// TIA Portal V15.1 export
// export: Created 2026-11-02T18:55:10.9093708Z, ExportSetting WithDefaults, DisplayName Totally Integrated Automation Portal, DisplayVersion V15.1, DisplayName TIA Portal Openness, DisplayVersion V15.1, DisplayName STEP 7 Professional, DisplayVersion V15.1, DisplayName WinCC Professional, DisplayVersion V15.1
FUNCTION_BLOCK "Scrubber"   // FB2, LAD
TITLE = Scrubber
{ S7_Optimized_Access := 'TRUE' }
VERSION : 0.1
// Gas scrubber, docs/التشغيل.md §1
// stored: AutoNumber false, IsIECCheckEnabled false, IsRetainMemResEnabled false, MemoryReserve 100, SetENOAutomatically False, UDAEnableTagReadback false
   VAR_INPUT
      PSH : Bool;   // PSH-101 healthy (contact closed)
      LSH : Bool;   // LSH-102 healthy
      LSHH : Bool;   // LSHH-103 healthy
      EStopOK : Bool;   // Sys.EStopOK
      ResetPulse : Bool;   // Sys.ResetPulse
      FirstScan : Bool;   // Sys.FirstScan
      TDrnOn : Time;   // Par.TDrnOn_V (C04)
      TDrnOff : Time;   // Par.TDrnOff_V (C04)
      TDrnMax : Time;   // Par.TDrnMax_V (C04a)
   END_VAR
   VAR_OUTPUT
      Tripped : Bool;   // Suction trip latch C01/C02/C03/C05: XV-403 closed until RESET
      FlareTrip : Bool;   // Flare trip latch C01/C02/C03: XV-401 open until RESET
      ValvesNormal : Bool;   // No trip latched: flare closed and suction open (HMI)
      FlareCmd : Bool;   // Q0.2 XV-401 (NO): 1 = energised = closed
      DrainCmd : Bool;   // Q0.3 XV-402 (NC): 1 = energised = open (C04 / C05)
      SuctionCmd : Bool;   // Q0.4 XV-403 (NC): 1 = energised = open
      F_DrainTO : Bool;   // C04a: drain open too long, latched until RESET
      F_LshFault : Bool;   // C04b: LSHH-103 without LSH-102, latched until RESET
      Alm_PSH : Bool;   // HMI alarm C03
      Alm_LSH : Bool;   // HMI alarm C04
      Alm_LSHH : Bool;   // HMI alarm C05
      Cause_EStop : Bool;   // C06a / F44: E-STOP cause, latched until healthy RESET
      Cause_PSH : Bool;   // C06a / F44: PSH-101 cause, latched until healthy RESET
      Cause_LSHH : Bool;   // C06a / F44: LSHH-103 cause, latched until healthy RESET
      Cause_PwrUp : Bool;   // C06a / F44: power-up cause, latched until healthy RESET
      FirstOut : Int;   // C06a / 0007 D5: 0 none, 1 E-STOP, 2 PSH, 3 LSHH, 4 power-up
   END_VAR
   VAR
      LevelHigh : Bool;
      DrnDemand : Bool;
      T_DrnOn : TON_TIME;
      T_DrnOff : TON_TIME;
      T_DrnMax : TON_TIME;
      T_LshFlt : TON_TIME;
   END_VAR
BEGIN

REGION Network 1: C04 — LSH-102 high level alarm
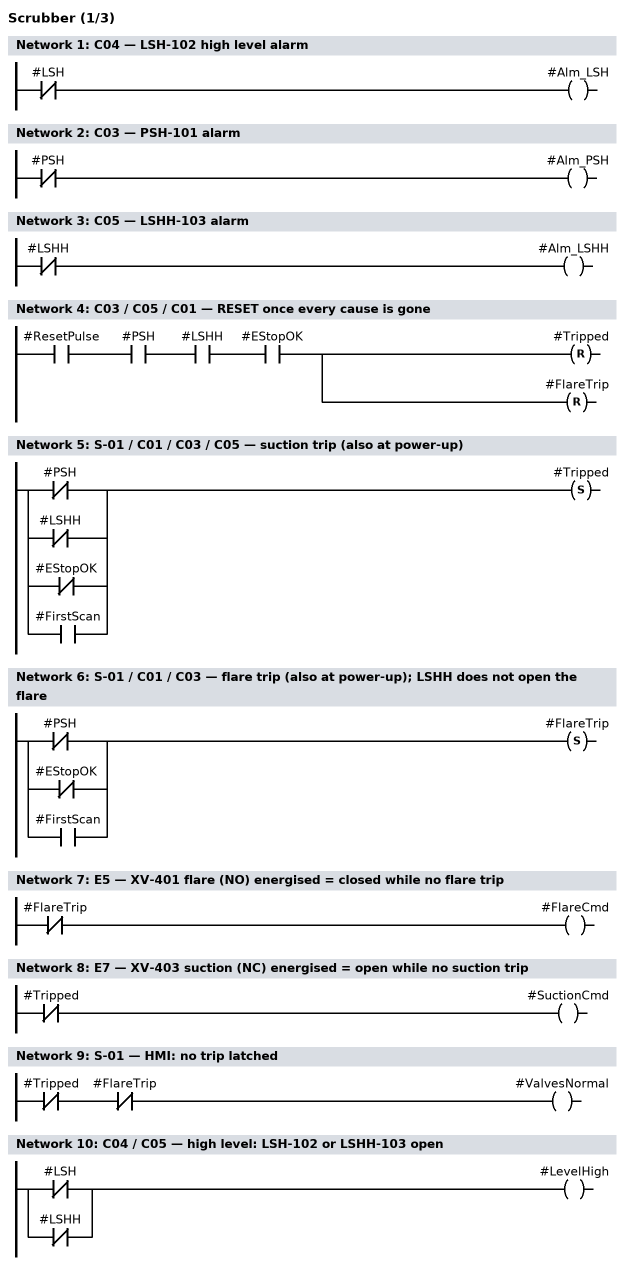
   RUNG wire#powerrail
      I_Contact( #LSH )
      Coil( #Alm_LSH )
   END_RUNG
   // the same network as SCL:
   #Alm_LSH := NOT #LSH;
END_REGION

REGION Network 2: C03 — PSH-101 alarm
   RUNG wire#powerrail
      I_Contact( #PSH )
      Coil( #Alm_PSH )
   END_RUNG
   // the same network as SCL:
   #Alm_PSH := NOT #PSH;
END_REGION

REGION Network 3: C05 — LSHH-103 alarm
   RUNG wire#powerrail
      I_Contact( #LSHH )
      Coil( #Alm_LSHH )
   END_RUNG
   // the same network as SCL:
   #Alm_LSHH := NOT #LSHH;
END_REGION

REGION Network 4: C03 / C05 / C01 — RESET once every cause is gone
   RUNG wire#powerrail
      Contact( #ResetPulse )
      Contact( #PSH )
      Contact( #LSHH )
      Contact( #EStopOK )
      wire#w1
      R_Coil( #Tripped )
   END_RUNG
   RUNG wire#w1
      R_Coil( #FlareTrip )
   END_RUNG
   // the same network as SCL:
   IF #ResetPulse AND #PSH AND #LSHH AND #EStopOK THEN
       #Tripped := FALSE;
       #FlareTrip := FALSE;
   END_IF;
END_REGION

REGION Network 5: S-01 / C01 / C03 / C05 — suction trip (also at power-up)
   RUNG wire#powerrail
      I_Contact( #PSH )
      wire#w1
      S_Coil( #Tripped )
   END_RUNG
   RUNG wire#powerrail
      I_Contact( #LSHH )
   END_RUNG wire#w1
   RUNG wire#powerrail
      I_Contact( #EStopOK )
   END_RUNG wire#w1
   RUNG wire#powerrail
      Contact( #FirstScan )
   END_RUNG wire#w1
   // the same network as SCL:
   IF NOT #PSH OR NOT #LSHH OR NOT #EStopOK OR #FirstScan THEN #Tripped := TRUE; END_IF;
END_REGION

REGION Network 6: S-01 / C01 / C03 — flare trip (also at power-up); LSHH does not open the flare
   RUNG wire#powerrail
      I_Contact( #PSH )
      wire#w1
      S_Coil( #FlareTrip )
   END_RUNG
   RUNG wire#powerrail
      I_Contact( #EStopOK )
   END_RUNG wire#w1
   RUNG wire#powerrail
      Contact( #FirstScan )
   END_RUNG wire#w1
   // the same network as SCL:
   IF NOT #PSH OR NOT #EStopOK OR #FirstScan THEN #FlareTrip := TRUE; END_IF;
END_REGION

REGION Network 7: E5 — XV-401 flare (NO) energised = closed while no flare trip
   RUNG wire#powerrail
      I_Contact( #FlareTrip )
      Coil( #FlareCmd )
   END_RUNG
   // the same network as SCL:
   #FlareCmd := NOT #FlareTrip;
END_REGION

REGION Network 8: E7 — XV-403 suction (NC) energised = open while no suction trip
   RUNG wire#powerrail
      I_Contact( #Tripped )
      Coil( #SuctionCmd )
   END_RUNG
   // the same network as SCL:
   #SuctionCmd := NOT #Tripped;
END_REGION

REGION Network 9: S-01 — HMI: no trip latched
   RUNG wire#powerrail
      I_Contact( #Tripped )
      I_Contact( #FlareTrip )
      Coil( #ValvesNormal )
   END_RUNG
   // the same network as SCL:
   #ValvesNormal := NOT #Tripped AND NOT #FlareTrip;
END_REGION

REGION Network 10: C04 / C05 — high level: LSH-102 or LSHH-103 open
   RUNG wire#powerrail
      I_Contact( #LSH )
      wire#w1
      Coil( #LevelHigh )
   END_RUNG
   RUNG wire#powerrail
      I_Contact( #LSHH )
   END_RUNG wire#w1
   // the same network as SCL:
   #LevelHigh := NOT #LSH OR NOT #LSHH;
END_REGION

REGION Network 11: C04 — drain demand after TDRN_ON of high level
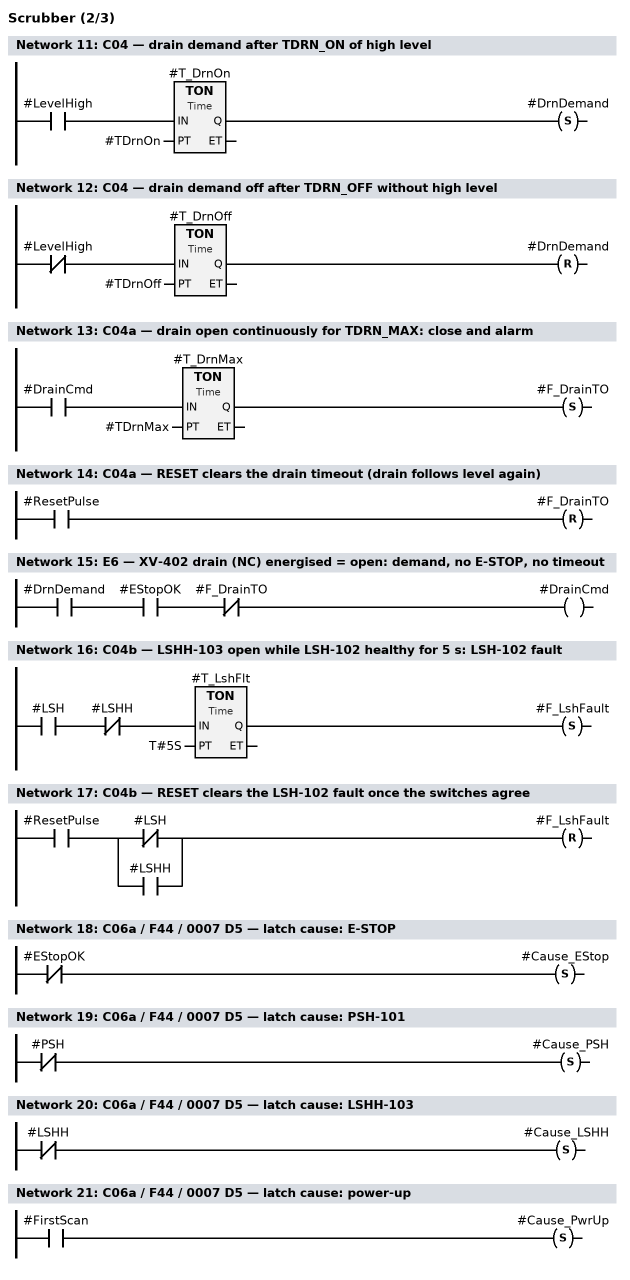
   RUNG wire#powerrail
      Contact( #LevelHigh )
      { S7_Templates := "time_type := Time" } #T_DrnOn.TON(pt := #TDrnOn, et =>)
      S_Coil( #DrnDemand )
   END_RUNG
   // the same network as SCL:
   #T_DrnOn(IN := #LevelHigh, PT := #TDrnOn);   // TON
   IF #T_DrnOn.Q THEN #DrnDemand := TRUE; END_IF;
END_REGION

REGION Network 12: C04 — drain demand off after TDRN_OFF without high level
   RUNG wire#powerrail
      I_Contact( #LevelHigh )
      { S7_Templates := "time_type := Time" } #T_DrnOff.TON(pt := #TDrnOff, et =>)
      R_Coil( #DrnDemand )
   END_RUNG
   // the same network as SCL:
   #T_DrnOff(IN := NOT #LevelHigh, PT := #TDrnOff);   // TON
   IF #T_DrnOff.Q THEN #DrnDemand := FALSE; END_IF;
END_REGION

REGION Network 13: C04a — drain open continuously for TDRN_MAX: close and alarm
   RUNG wire#powerrail
      Contact( #DrainCmd )
      { S7_Templates := "time_type := Time" } #T_DrnMax.TON(pt := #TDrnMax, et =>)
      S_Coil( #F_DrainTO )
   END_RUNG
   // the same network as SCL:
   #T_DrnMax(IN := #DrainCmd, PT := #TDrnMax);   // TON
   IF #T_DrnMax.Q THEN #F_DrainTO := TRUE; END_IF;
END_REGION

REGION Network 14: C04a — RESET clears the drain timeout (drain follows level again)
   RUNG wire#powerrail
      Contact( #ResetPulse )
      R_Coil( #F_DrainTO )
   END_RUNG
   // the same network as SCL:
   IF #ResetPulse THEN #F_DrainTO := FALSE; END_IF;
END_REGION

REGION Network 15: E6 — XV-402 drain (NC) energised = open: demand, no E-STOP, no timeout
   RUNG wire#powerrail
      Contact( #DrnDemand )
      Contact( #EStopOK )
      I_Contact( #F_DrainTO )
      Coil( #DrainCmd )
   END_RUNG
   // the same network as SCL:
   #DrainCmd := #DrnDemand AND #EStopOK AND NOT #F_DrainTO;
END_REGION

REGION Network 16: C04b — LSHH-103 open while LSH-102 healthy for 5 s: LSH-102 fault
   RUNG wire#powerrail
      Contact( #LSH )
      I_Contact( #LSHH )
      { S7_Templates := "time_type := Time" } #T_LshFlt.TON(pt := T#5S, et =>)
      S_Coil( #F_LshFault )
   END_RUNG
   // the same network as SCL:
   #T_LshFlt(IN := #LSH AND NOT #LSHH, PT := T#5S);   // TON
   IF #T_LshFlt.Q THEN #F_LshFault := TRUE; END_IF;
END_REGION

REGION Network 17: C04b — RESET clears the LSH-102 fault once the switches agree
   RUNG wire#powerrail
      Contact( #ResetPulse )
      wire#w1
      I_Contact( #LSH )
      wire#w2
      R_Coil( #F_LshFault )
   END_RUNG
   RUNG wire#w1
      Contact( #LSHH )
   END_RUNG wire#w2
   // the same network as SCL:
   IF #ResetPulse AND (NOT #LSH OR #LSHH) THEN #F_LshFault := FALSE; END_IF;
END_REGION

REGION Network 18: C06a / F44 / 0007 D5 — latch cause: E-STOP
   RUNG wire#powerrail
      I_Contact( #EStopOK )
      S_Coil( #Cause_EStop )
   END_RUNG
   // the same network as SCL:
   IF NOT #EStopOK THEN #Cause_EStop := TRUE; END_IF;
END_REGION

REGION Network 19: C06a / F44 / 0007 D5 — latch cause: PSH-101
   RUNG wire#powerrail
      I_Contact( #PSH )
      S_Coil( #Cause_PSH )
   END_RUNG
   // the same network as SCL:
   IF NOT #PSH THEN #Cause_PSH := TRUE; END_IF;
END_REGION

REGION Network 20: C06a / F44 / 0007 D5 — latch cause: LSHH-103
   RUNG wire#powerrail
      I_Contact( #LSHH )
      S_Coil( #Cause_LSHH )
   END_RUNG
   // the same network as SCL:
   IF NOT #LSHH THEN #Cause_LSHH := TRUE; END_IF;
END_REGION

REGION Network 21: C06a / F44 / 0007 D5 — latch cause: power-up
   RUNG wire#powerrail
      Contact( #FirstScan )
      S_Coil( #Cause_PwrUp )
   END_RUNG
   // the same network as SCL:
   IF #FirstScan THEN #Cause_PwrUp := TRUE; END_IF;
END_REGION

REGION Network 22: C06a / F44 / 0007 D5 — first-out 1: E-STOP (only if none)
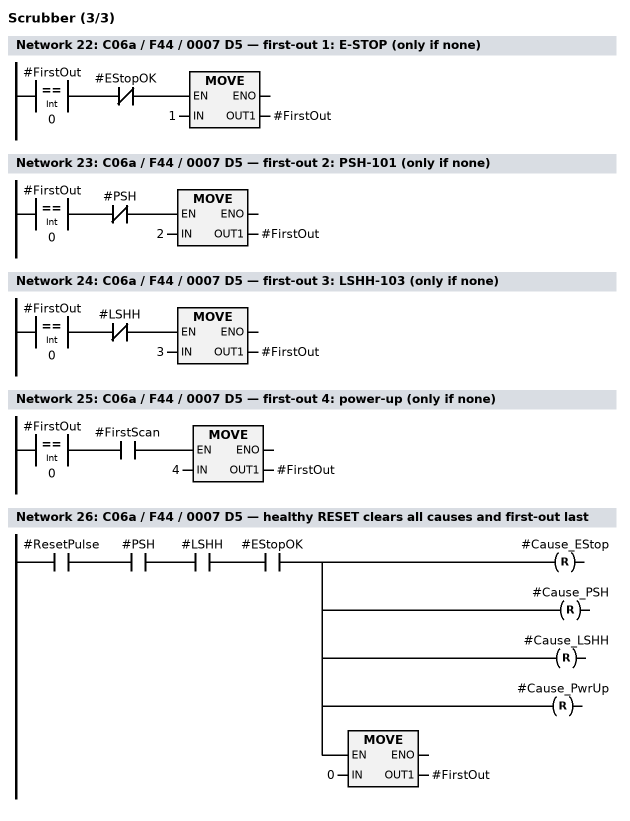
   RUNG wire#powerrail
      { S7_Templates := "SrcType := Int" } EQ_Contact(in1 := #FirstOut, in2 := 0)
      I_Contact( #EStopOK )
      { S7_GenerateENO := "TRUE" } Move(in := 1, out1 => #FirstOut)
   END_RUNG
   // the same network as SCL:
   IF (#FirstOut = 0) AND NOT #EStopOK THEN #FirstOut := 1; END_IF;
END_REGION

REGION Network 23: C06a / F44 / 0007 D5 — first-out 2: PSH-101 (only if none)
   RUNG wire#powerrail
      { S7_Templates := "SrcType := Int" } EQ_Contact(in1 := #FirstOut, in2 := 0)
      I_Contact( #PSH )
      { S7_GenerateENO := "TRUE" } Move(in := 2, out1 => #FirstOut)
   END_RUNG
   // the same network as SCL:
   IF (#FirstOut = 0) AND NOT #PSH THEN #FirstOut := 2; END_IF;
END_REGION

REGION Network 24: C06a / F44 / 0007 D5 — first-out 3: LSHH-103 (only if none)
   RUNG wire#powerrail
      { S7_Templates := "SrcType := Int" } EQ_Contact(in1 := #FirstOut, in2 := 0)
      I_Contact( #LSHH )
      { S7_GenerateENO := "TRUE" } Move(in := 3, out1 => #FirstOut)
   END_RUNG
   // the same network as SCL:
   IF (#FirstOut = 0) AND NOT #LSHH THEN #FirstOut := 3; END_IF;
END_REGION

REGION Network 25: C06a / F44 / 0007 D5 — first-out 4: power-up (only if none)
   RUNG wire#powerrail
      { S7_Templates := "SrcType := Int" } EQ_Contact(in1 := #FirstOut, in2 := 0)
      Contact( #FirstScan )
      { S7_GenerateENO := "TRUE" } Move(in := 4, out1 => #FirstOut)
   END_RUNG
   // the same network as SCL:
   IF (#FirstOut = 0) AND #FirstScan THEN #FirstOut := 4; END_IF;
END_REGION

REGION Network 26: C06a / F44 / 0007 D5 — healthy RESET clears all causes and first-out last
   RUNG wire#powerrail
      Contact( #ResetPulse )
      Contact( #PSH )
      Contact( #LSHH )
      Contact( #EStopOK )
      wire#w1
      R_Coil( #Cause_EStop )
   END_RUNG
   RUNG wire#w1
      R_Coil( #Cause_PSH )
   END_RUNG
   RUNG wire#w1
      R_Coil( #Cause_LSHH )
   END_RUNG
   RUNG wire#w1
      R_Coil( #Cause_PwrUp )
   END_RUNG
   RUNG wire#w1
      { S7_GenerateENO := "TRUE" } Move(in := 0, out1 => #FirstOut)
   END_RUNG
   // the same network as SCL:
   IF #ResetPulse AND #PSH AND #LSHH AND #EStopOK THEN
       #Cause_EStop := FALSE;
       #Cause_PSH := FALSE;
       #Cause_LSHH := FALSE;
       #Cause_PwrUp := FALSE;
       #FirstOut := 0;
   END_IF;
END_REGION
END_FUNCTION_BLOCK
